Staubli VAL3: getProgItemSize.pgx

public program getProgItemSize(string x_sKey, num& x_nSize)
begin
  x_nSize=size(progTemp:pProgItem[x_sKey].pProgTemplate)
end
